// TIA Portal V21 export
// export: Created 2026-10-12T11:32:14.0782283Z, ExportSetting WithDefaults, DisplayName Totally Integrated Automation Portal, DisplayVersion V21, DisplayName STEP 7 Professional, DisplayVersion V21, DisplayName STEP 7 Safety, DisplayVersion V21, DisplayName Tech WebApplication, DisplayVersion V21, DisplayName WinCC Basic/Comfort/Advanced, DisplayVersion V21, DisplayName WinCC Unified, DisplayVersion V21
FUNCTION "FC_MANUAL" : Void   // FC2, LAD
{ S7_Optimized_Access := 'TRUE' }
VERSION : 0.1
// stored: AutoNumber true, IsIECCheckEnabled false, SetENOAutomatically false, UDAEnableTagReadback false
   VAR_TEMP   // added for the SCL form of the ladder/FBD networks
      _w1 : Bool;
   END_VAR
BEGIN

REGION Network 1: MOTOR FWD /REV ON
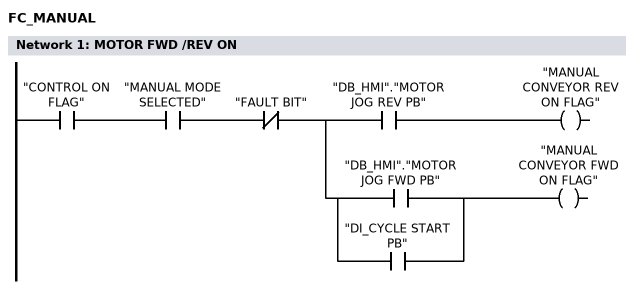
   RUNG wire#powerrail
      Contact( "CONTROL ON FLAG" )
      Contact( "MANUAL MODE SELECTED" )
      I_Contact( "FAULT BIT" )
      wire#w1
      Contact( "DB_HMI"."MOTOR JOG REV PB" )
      Coil( "MANUAL CONVEYOR REV ON FLAG" )
   END_RUNG
   RUNG wire#w1
      Contact( "DB_HMI"."MOTOR JOG FWD PB" )
      wire#w2
      Coil( "MANUAL CONVEYOR FWD ON FLAG" )
   END_RUNG
   RUNG wire#w1
      Contact( "DI_CYCLE START PB" )
   END_RUNG wire#w2
   // the same network as SCL:
   #_w1 := "CONTROL ON FLAG" AND "MANUAL MODE SELECTED" AND NOT "FAULT BIT";
   "MANUAL CONVEYOR REV ON FLAG" := #_w1 AND "DB_HMI"."MOTOR JOG REV PB";
   "MANUAL CONVEYOR FWD ON FLAG" := #_w1 AND ("DB_HMI"."MOTOR JOG FWD PB" OR "DI_CYCLE START PB");
END_REGION
END_FUNCTION
